(* IEC 61131-3 sources: matiec/tests/warnings, 3 files *)

(* ---- ok_extensible_functions.st ---- *)
(* Calls of extensible standard functions. Their extensible operands are passed
   through a C "...", so they undergo default argument promotions: REAL ones
   become double, triggering -Wdouble-promotion, and va_start() must not take
   such an operand as its last named parameter (clang's -Wvarargs).
   Calls come from ST, from IL, and from the inline functions that get ENO. *)

FUNCTION_BLOCK fb_il
  VAR_INPUT
    ra, rb : REAL;
  END_VAR
  VAR_OUTPUT
    rmax, rmax2 : REAL;
    smax : SINT;
    ra_gt_rb : BOOL;
  END_VAR
  VAR
    sa : SINT;
  END_VAR
  LD ra
  MAX rb, 1.5
  ST rmax
  MAX(
    IN1 := ra,
    IN2 := rb
  )
  ST rmax2
  LD sa
  MAX 3
  ST smax
  LD ra
  GT rb
  ST ra_gt_rb
END_FUNCTION_BLOCK

PROGRAM program0
  VAR
    sa, sb : SINT;
    ra, rb, rc : REAL;
    ba, bb : BOOL;
    ta, tb : TIME;
    stra, strb : STRING;
    k : INT;
    ok : BOOL;
    il : fb_il;
  END_VAR

  rc := ADD(ra, rb, 2.5);
  rc := MAX(ra, rb);
  rc := MUX(k, ra, rb, rc);
  sa := MUL(sa, sb, 3);
  ba := XOR(ba, bb, TRUE);
  ba := GT(ra, rb, rc);
  ba := EQ(ta, tb);
  stra := CONCAT(stra, strb, 'x');
  rc := ADD(EN := ba, IN1 := ra, IN2 := rb, ENO => ok);
  sa := MAX(EN := ba, IN1 := sa, IN2 := sb, ENO => ok);
  il(ra := ra, rb := rb);
END_PROGRAM

CONFIGURATION config
  RESOURCE resource1 ON PLC
    TASK main_task(INTERVAL := T#1000ms, PRIORITY := 0);
    PROGRAM instance0 WITH main_task : program0;
  END_RESOURCE
END_CONFIGURATION

(* ---- ok_resource_globals.st ---- *)
(* Globals of resources, that POUs use as VAR_EXTERNAL, as in Beremiz's
   first_steps example. Their getters (__GET_GLOBAL_<name>) are defined in the
   C file of each resource only, while config.c also includes POUS.c, for the
   constructors of POUs. So do calls to functions with VAR_OUTPUT, that are
   made through inline wrappers. *)

FUNCTION double_it : DINT
  VAR_INPUT
    i : DINT;
  END_VAR
  VAR_OUTPUT
    o : DINT;
  END_VAR
  o := i * 2;
  double_it := o;
END_FUNCTION

FUNCTION_BLOCK fb0
  VAR_EXTERNAL
    resource_global : DINT;
  END_VAR
  VAR
    doubled : DINT;
  END_VAR
  resource_global := double_it(i := resource_global, o => doubled);
END_FUNCTION_BLOCK

PROGRAM program0
  VAR_EXTERNAL
    resource_global : DINT;
    resource_timer : TON;
  END_VAR
  VAR
    fb_instance : fb0;
    doubled : DINT;
  END_VAR
  resource_timer(IN := TRUE, PT := T#1s);
  fb_instance();
  resource_global := double_it(i := resource_global, o => doubled);
END_PROGRAM

CONFIGURATION config
  RESOURCE resource1 ON PLC
    VAR_GLOBAL
      resource_global : DINT := 1;
      resource_timer : TON;
    END_VAR
    TASK main_task(INTERVAL := T#1000ms, PRIORITY := 0);
    PROGRAM instance0 WITH main_task : program0;
  END_RESOURCE
  RESOURCE resource2 ON PLC
    VAR_GLOBAL
      resource_global : DINT := 2;
      resource_timer : TON;
    END_VAR
    TASK main_task(INTERVAL := T#20ms, PRIORITY := 0);
    PROGRAM instance1 WITH main_task : program0;
  END_RESOURCE
END_CONFIGURATION

(* ---- ok_conditions.st ---- *)
(* Conditions of IF, ELSIF, WHILE and CASE that compare a variable with '='.
   They become C if and while statements, that put their condition in
   parentheses, and clang warns about "if ((a == b))" (-Wparentheses-equality). *)

PROGRAM program0
  VAR
    ia : INT;
  END_VAR

  IF ia = 5 THEN
    ia := 0;
  ELSIF ia = 6 THEN
    ia := 1;
  END_IF;
  WHILE ia = 7 DO
    ia := 8;
  END_WHILE;
  CASE ia OF
    1: ia := 2;
    3, 4..5: ia := 6;
  END_CASE;
END_PROGRAM

CONFIGURATION config
  RESOURCE resource1 ON PLC
    TASK main_task(INTERVAL := T#1000ms, PRIORITY := 0);
    PROGRAM instance0 WITH main_task : program0;
  END_RESOURCE
END_CONFIGURATION
